FUNCTION_BLOCK basicEEEBruto (* Logica unica da elevatoria de esgoto bruto (3 bombas, 2 operando + 1 reserva) *)
  (* Standard: 61499-2 *)
  (* Version 1.6, 21/10/2026, Hidryco, Hidryco, 1.6: PID de nivel em Hz (minimo, maximo, preset e saida; 60 Hz = 100 %); STS_VELOCIDADE da IHM em Hz. 1.5: faixas da necessidade pela % da altura do poco (nivPct); stsNivel (IHM) continua em metros. 1.4: IHM: nivel, saida do PID, velocidade e tempo restante no maximo 1 vez por segundo (TICK). 1.3: pressao L/LL do PIT-01 inibida com as bombas paradas mesmo com cfgTempoPartidaPressao = 0. 1.2: emergencia do PCM NF. 1.1: emergencia do painel e falha de comunicacao dos ATV630. 1.0: faixas de nivel, revezamento por tempo, PID de velocidade, HH do Nereda, operacao pelas boias, falha de recalque *)
  PACKAGE Hidryco.HidrycoLib;
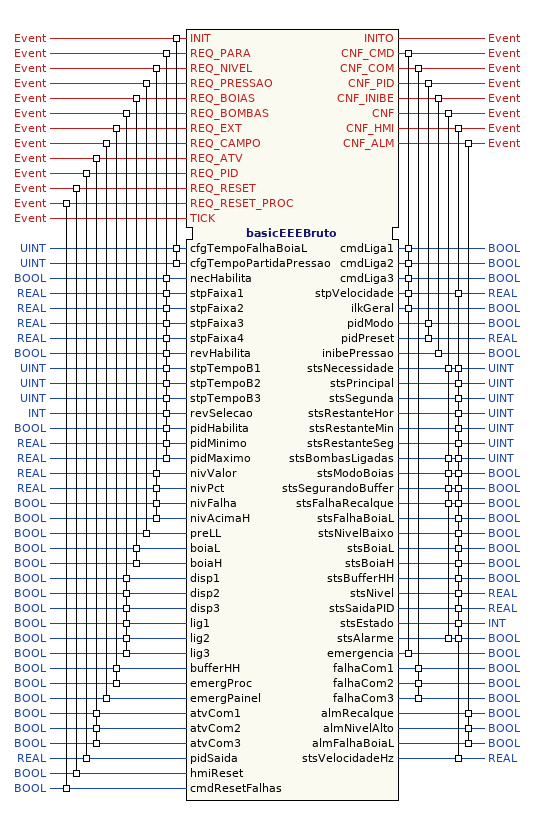
  EVENT_INPUT
    INIT WITH cfgTempoFalhaBoiaL, cfgTempoPartidaPressao; (* Inicializacao *)
    REQ_PARA WITH necHabilita, stpFaixa1, stpFaixa2, stpFaixa3, stpFaixa4, revHabilita, stpTempoB1, stpTempoB2, stpTempoB3, revSelecao, pidHabilita, pidMinimo, pidMaximo; (* Parametros da IHM (persistentes) *)
    REQ_NIVEL WITH nivValor, nivPct, nivFalha, nivAcimaH; (* LIT-03 *)
    REQ_PRESSAO WITH preLL; (* PIT-01 *)
    REQ_BOIAS WITH boiaL, boiaH; (* Boias *)
    REQ_BOMBAS WITH disp1, disp2, disp3, lig1, lig2, lig3; (* Estado das bombas *)
    REQ_EXT WITH bufferHH, emergProc; (* Processo *)
    REQ_CAMPO WITH emergPainel; (* Emergencia do painel *)
    REQ_ATV WITH atvCom1, atvCom2, atvCom3; (* Comunicacao dos ATV630 *)
    REQ_PID WITH pidSaida; (* Saida do PID *)
    REQ_RESET WITH hmiReset; (* Reset pela IHM *)
    REQ_RESET_PROC WITH cmdResetFalhas; (* Reset pelo processo *)
    TICK; (* Base de tempo de 1 s (E_CYCLE) *)
  END_EVENT
  EVENT_OUTPUT
    INITO; (* Inicializacao concluida *)
    CNF_CMD WITH cmdLiga1, cmdLiga2, cmdLiga3, stpVelocidade, ilkGeral, emergencia; (* Comandos para as bombas (na mudanca) *)
    CNF_COM WITH falhaCom1, falhaCom2, falhaCom3; (* Falha de comunicacao dos ATV630 para os motores (na mudanca e a cada leitura) *)
    CNF_PID WITH pidModo, pidPreset; (* Modo do pidCtl (na mudanca) *)
    CNF_INIBE WITH inibePressao; (* Inibicao dos alarmes baixos do PIT-01 (na mudanca) *)
    CNF WITH stsNecessidade, stsBombasLigadas, stsSegurandoBuffer, stsModoBoias, stsFalhaRecalque, stsAlarme; (* Status para o processo (na mudanca) *)
    CNF_HMI WITH stsNecessidade, stsPrincipal, stsSegunda, stsRestanteHor, stsRestanteMin, stsRestanteSeg, stsBombasLigadas, stsModoBoias, stsSegurandoBuffer, stsFalhaRecalque, stsFalhaBoiaL, stsNivelBaixo, stsBoiaL, stsBoiaH, stsBufferHH, stsNivel, stsSaidaPID, stpVelocidade, stsEstado, stsAlarme, stsVelocidadeHz; (* Status para a IHM (na mudanca) *)
    CNF_ALM WITH almRecalque, almNivelAlto, almFalhaBoiaL; (* Alarmes para os ALARM_BIT (na mudanca) *)
  END_EVENT
  VAR_INPUT
    cfgTempoFalhaBoiaL : UINT := 10; (* Operacao pelas boias com a boia LSL com defeito: bombas ficam ligadas este tempo (min) depois que a LSH desce *)
    cfgTempoPartidaPressao : UINT := 30; (* Alarmes L/LL do PIT-01 inibidos ate a bomba estar ligada ha este tempo (s); tambem inibidos com as bombas paradas *)
    necHabilita : BOOL; (* IHM: automatico da elevatoria habilitado (NEC_CMD_HABILITA) *)
    stpFaixa1 : REAL; (* IHM: com 1 bomba, desliga abaixo deste nivel (STP_LIMITE_FAIXA_1) *)
    stpFaixa2 : REAL; (* IHM: com 2 bombas, desliga a 2a abaixo deste nivel (STP_LIMITE_FAIXA_2) *)
    stpFaixa3 : REAL; (* IHM: parada, liga a 1a bomba neste nivel (STP_LIMITE_FAIXA_3) *)
    stpFaixa4 : REAL; (* IHM: com 1 bomba, liga a 2a neste nivel (STP_LIMITE_FAIXA_4) *)
    revHabilita : BOOL; (* IHM: revezamento por tempo habilitado (REV_CMD_HABILITA) *)
    stpTempoB1 : UINT; (* IHM: horas da bomba 1 como principal antes da troca; 0 = sem troca por tempo (STP_TEMPO_B1) *)
    stpTempoB2 : UINT; (* IHM: horas da bomba 2 como principal antes da troca; 0 = sem troca por tempo (STP_TEMPO_B2) *)
    stpTempoB3 : UINT; (* IHM: horas da bomba 3 como principal antes da troca; 0 = sem troca por tempo (STP_TEMPO_B3) *)
    revSelecao : INT; (* IHM: bomba principal 1, 2 ou 3 (CMD_SELECAO_BOMBA); comeca por ela ao escolher e a cada nova partida *)
    pidHabilita : BOOL; (* IHM: velocidade pelo PID de nivel (PID_CMD_HABILITA); FALSE = velocidade maxima *)
    pidMinimo : REAL; (* IHM: velocidade minima / saida minima do PID, % (STP_MINIMO) *)
    pidMaximo : REAL; (* IHM: velocidade maxima / saida maxima do PID, % (STP_MAXIMO) *)
    nivValor : REAL; (* LIT-03: nivel (unidade de engenharia) *)
    nivPct : REAL; (* LIT-03: nivel em % da altura do poco (faixas da necessidade) *)
    nivFalha : BOOL; (* LIT-03: sinal em falha agora *)
    nivAcimaH : BOOL; (* LIT-03: nivel acima do setpoint H agora (alarme H habilitado) *)
    preLL : BOOL; (* PIT-01: alarme LL de pressao (ja com o tempo do sensor) *)
    boiaL : BOOL; (* LSL-04: TRUE = boia levantada (nivel acima do baixo) *)
    boiaH : BOOL; (* LSH-05: TRUE = boia levantada (nivel alto) *)
    disp1 : BOOL; (* Bomba 1 disponivel para o automatico *)
    disp2 : BOOL; (* Bomba 2 disponivel para o automatico *)
    disp3 : BOOL; (* Bomba 3 disponivel para o automatico *)
    lig1 : BOOL; (* Bomba 1 ligada *)
    lig2 : BOOL; (* Bomba 2 ligada *)
    lig3 : BOOL; (* Bomba 3 ligada *)
    bufferHH : BOOL; (* Processo: nivel HH do tanque de equalizacao do Nereda (40-LT-0001) *)
    emergProc : BOOL; (* Processo: emergencia (entrada stsEmergencia do CAT) *)
    emergPainel : BOOL; (* Campo: emergencia do PCM EEE Bruto, NF (TRUE = normal; FALSE = em emergencia) *)
    atvCom1 : BOOL; (* ATV630 da bomba 1: comunicacao ativa (ComStatus do HW CAT) *)
    atvCom2 : BOOL; (* ATV630 da bomba 2: comunicacao ativa (ComStatus do HW CAT) *)
    atvCom3 : BOOL; (* ATV630 da bomba 3: comunicacao ativa (ComStatus do HW CAT) *)
    pidSaida : REAL; (* Saida do pidCtl (%) *)
    hmiReset : BOOL; (* IHM: reset *)
    cmdResetFalhas : BOOL; (* Processo: reset (com E_RESET_FALHAS) *)
  END_VAR
  VAR_OUTPUT
    cmdLiga1 : BOOL; (* Comando automatico da bomba 1 *)
    cmdLiga2 : BOOL; (* Comando automatico da bomba 2 *)
    cmdLiga3 : BOOL; (* Comando automatico da bomba 3 *)
    stpVelocidade : REAL; (* Velocidade das bombas ligadas (%) *)
    ilkGeral : BOOL; (* Intertravamento geral das bombas (LSL em nivel baixo ou falha de recalque); vale em qualquer modo *)
    pidModo : BOOL; (* pidCtl em automatico *)
    pidPreset : REAL; (* Valor do pidCtl em manual (%) *)
    inibePressao : BOOL; (* Inibe os alarmes L/LL do PIT-01 *)
    stsNecessidade : UINT; (* Numero de bombas pedidas (0, 1, 2) *)
    stsPrincipal : UINT; (* Bomba principal (1..3) *)
    stsSegunda : UINT; (* Bomba que entra como 2a (0 = nenhuma disponivel) *)
    stsRestanteHor : UINT; (* Tempo para a troca da principal (h) *)
    stsRestanteMin : UINT; (* Tempo para a troca da principal (min) *)
    stsRestanteSeg : UINT; (* Tempo para a troca da principal (s) *)
    stsBombasLigadas : UINT; (* Bombas ligadas *)
    stsModoBoias : BOOL; (* Operacao de emergencia pelas boias (LIT-03 em falha) *)
    stsSegurandoBuffer : BOOL; (* Elevatoria parada segurando o esgoto (HH do tanque do Nereda) *)
    stsFalhaRecalque : BOOL; (* Falha de recalque (pressao LL com bomba ligada) - memorizada ate o reset *)
    stsFalhaBoiaL : BOOL; (* Boia LSL com defeito (LSH levantada com a LSL abaixada) - memorizada ate o reset *)
    stsNivelBaixo : BOOL; (* LSL em nivel baixo: bombas intertravadas *)
    stsBoiaL : BOOL; (* LSL-04 *)
    stsBoiaH : BOOL; (* LSH-05 *)
    stsBufferHH : BOOL; (* HH do tanque do Nereda *)
    stsNivel : REAL; (* Nivel do poco *)
    stsSaidaPID : REAL; (* Saida do PID (%) *)
    stsEstado : INT; (* 0 parada, 1 bombeando, 2 segurando (HH Nereda), 3 pelas boias, 4 falha de recalque, 5 nivel baixo (LSL), 6 automatico desabilitado, 7 emergencia *)
    stsAlarme : BOOL; (* Algum alarme da elevatoria *)
    emergencia : BOOL; (* Emergencia para as bombas (painel OU processo) *)
    falhaCom1 : BOOL; (* Falha de comunicacao com o ATV630 da bomba 1 (publicada no stsFalhaComunicacao do motor) *)
    falhaCom2 : BOOL; (* Falha de comunicacao com o ATV630 da bomba 2 (publicada no stsFalhaComunicacao do motor) *)
    falhaCom3 : BOOL; (* Falha de comunicacao com o ATV630 da bomba 3 (publicada no stsFalhaComunicacao do motor) *)
    almRecalque : BOOL; (* ALARM_BIT falha de recalque *)
    almNivelAlto : BOOL; (* ALARM_BIT nivel alto (LSH) *)
    almFalhaBoiaL : BOOL; (* ALARM_BIT defeito da boia LSL *)
    stsVelocidadeHz : REAL; (* Velocidade enviada as bombas em Hz (IHM/SCADA) *)
  END_VAR
  VAR
    initDone : BOOL;
    initPass : BOOL;
    bReset : BOOL;
    bNivelRecebido : BOOL; (* Ja houve leitura do LIT-03 *)
    bBoiasRecebidas : BOOL; (* Ja houve leitura das boias *)
    bNivelOk : BOOL; (* LIT-03 valido *)
    bAlgumaLigada : BOOL;
    bLiberadoHH : BOOL; (* HH do Nereda: liberado pelo nivel H do poco *)
    iNec : UINT; (* Numero de bombas pedidas *)
    oldNec : UINT;
    bCampoRecebido : BOOL; (* Ja houve leitura da emergencia do painel *)
    iPrincipal : UINT := 1; (* Bomba principal (revezamento) *)
    iSel : INT; (* Selecao da principal valida (1..3) *)
    oldSel : INT; (* Ultima selecao aplicada *)
    iUso : UINT; (* Principal em uso (fixa indisponivel = proxima) *)
    iSeg : UINT; (* 2a bomba *)
    iProx : UINT;
    iCand : UINT;
    i : UINT;
    bDisp : BOOL;
    bDispP : BOOL;
    bLigP : BOOL;
    uSegPrincipal : UDINT; (* Segundos da principal ligada desde a ultima troca *)
    uLimite : UDINT;
    uResta : UDINT;
    uTempoBoia : UDINT; (* Contagem (s) da operacao pelas boias com a LSL com defeito *)
    uSegLigada : UDINT; (* Segundos com bomba ligada (inibicao do PIT-01) *)
    wCmd : WORD;
    oldCmd : WORD := 16#FFFF;
    oldVel : REAL := -1.0;
    oldPidModo : BOOL;
    oldPreset : REAL := -1.0;
    oldInibe : BOOL;
    wSts : WORD;
    oldSts : WORD := 16#FFFF;
    wHmi : WORD;
    oldHmi : WORD := 16#FFFF;
    oldNivel : REAL := -1.0;
    oldSaida : REAL := -1.0;
    oldResta : UDINT := 16#FFFFFFFF;
    hmiVel : REAL := -1.0;
    oldEstado : INT := -1;
    oldInfo : UINT := 16#FFFF;
    uInfo : UINT;
    wAlm : WORD;
    oldAlm : WORD := 16#FFFF;
    wCom : WORD;
    oldCom : WORD := 16#FFFF;
  END_VAR
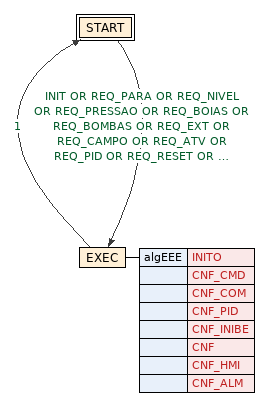
  EC_STATES
    START; (* Estado inicial *)
    EXEC : algEEE -> INITO, -> CNF_CMD, -> CNF_COM, -> CNF_PID, -> CNF_INIBE, -> CNF, -> CNF_HMI, -> CNF_ALM; (* Executa a logica; o algoritmo decide quais eventos saem *)
  END_STATES
  EC_TRANSITIONS
    START TO EXEC := INIT OR REQ_PARA OR REQ_NIVEL OR REQ_PRESSAO OR REQ_BOIAS OR REQ_BOMBAS OR REQ_EXT OR REQ_CAMPO OR REQ_ATV OR REQ_PID OR REQ_RESET OR REQ_RESET_PROC OR TICK;
    EXEC TO START := 1;
  END_TRANSITIONS
  ALGORITHM algEEE IN ST: (* Logica completa da elevatoria (um unico algoritmo) *)
(* =====================================================================
   basicEEEBruto v1.1 - Elevatoria de Esgoto Bruto (100-BS-01/02/03)
   Padrao das bibliotecas Schneider: eventos de saida desligados no inicio e
   ligados so na mudanca; tempos contados pelo TICK de 1 s (E_CYCLE do CAT).
   Regras (definidas pelo usuario, out/2026):
   - numero de bombas por faixas de nivel do LIT-03 (mesmas tags do CAT
     Necessidade_2_Equipamentos), no maximo 2; velocidade pelo PID de nivel;
   - revezamento: a principal selecionada (1, 2 ou 3) e a primeira a partir
     (ao escolher e sempre que as bombas partem de novo); com o revezamento
     habilitado troca apos STP_TEMPO_Bx horas ligada, na sequencia 1-2-3
     pulando a indisponivel; a 2a e a proxima da sequencia; principal
     indisponivel = troca na hora (tags do Revezamento_3_Motores);
   - HH do tanque do Nereda: a elevatoria para e segura o esgoto; volta a
     bombear quando o poco chega ao H dele (ou na LSH) - o tanque do Nereda
     tem extravasor; depois que esvazia ate a faixa 1, volta a segurar;
   - LIT-03 em falha: operacao pelas boias (LSH liga as 2 bombas na
     velocidade maxima; desligam quando a LSL abaixa; com a LSL com defeito,
     ficam cfgTempoFalhaBoiaL min depois que a LSH desce);
   - LSL abaixada desliga as bombas (ilkGeral) e elas voltam sozinhas;
   - PIT-01 em LL com bomba ligada = falha de recalque: para todas, alarma,
     memoriza ate o reset; L/LL do PIT-01 inibidos com as bombas paradas e
     nos primeiros cfgTempoPartidaPressao s depois da partida;
   - LSH so alarma (fora a operacao pelas boias e a liberacao do HH).
   v1.2: emergencia do PCM e NF (FALSE = em emergencia), so vale depois da
         1a leitura do campo.
   v1.1: emergencia do painel (campo) OU do processo vai para as bombas;
   falha de comunicacao de cada ATV630 = NOT ComStatus, publicada no
   stsFalhaComunicacao do motor (sem leitura = falha).
   ===================================================================== *)

(* ---- 0. Eventos de saida: so sai o que for ligado abaixo ---- *)
INITO     := FALSE;
CNF_CMD   := FALSE;
CNF_PID   := FALSE;
CNF_INIBE := FALSE;
CNF       := FALSE;
CNF_HMI   := FALSE;
CNF_ALM   := FALSE;
CNF_COM   := FALSE;

IF REQ_NIVEL THEN
    bNivelRecebido := TRUE;
END_IF;
IF REQ_BOIAS THEN
    bBoiasRecebidas := TRUE;
END_IF;
IF REQ_CAMPO THEN
    bCampoRecebido := TRUE;
END_IF;

(* ---- 1. Inicializacao ---- *)
IF INIT THEN
    initDone := TRUE;
    initPass := TRUE;
    INITO    := TRUE;
END_IF;
IF NOT initDone THEN
    RETURN;
END_IF;

bReset := (REQ_RESET AND hmiReset) OR (REQ_RESET_PROC AND cmdResetFalhas);
bAlgumaLigada := lig1 OR lig2 OR lig3;
stsBombasLigadas := 0;
IF lig1 THEN stsBombasLigadas := stsBombasLigadas + 1; END_IF;
IF lig2 THEN stsBombasLigadas := stsBombasLigadas + 1; END_IF;
IF lig3 THEN stsBombasLigadas := stsBombasLigadas + 1; END_IF;

(* ---- 2. Boias ---- *)
IF boiaH AND NOT boiaL THEN
    stsFalhaBoiaL := TRUE;                 (* LSH levantada com a LSL abaixada: LSL com defeito *)
END_IF;
IF bReset AND boiaL THEN
    stsFalhaBoiaL := FALSE;
END_IF;
(* nivel baixo: LSL abaixada (so se a LSL estiver confiavel); antes da 1a leitura, bloqueado *)
stsNivelBaixo := NOT bBoiasRecebidas OR (NOT boiaL AND NOT stsFalhaBoiaL);

(* ---- 3. Falha de recalque (PIT-01) ---- *)
IF bAlgumaLigada THEN
    IF TICK AND uSegLigada < UINT_TO_UDINT(cfgTempoPartidaPressao) THEN
        uSegLigada := uSegLigada + 1;
    END_IF;
ELSE
    uSegLigada := 0;
END_IF;
inibePressao := NOT bAlgumaLigada OR uSegLigada < UINT_TO_UDINT(cfgTempoPartidaPressao);   (* parada: inibido mesmo com o tempo = 0 *)
IF preLL AND NOT inibePressao THEN
    stsFalhaRecalque := TRUE;              (* pressao LL com bomba ligada: para todas *)
END_IF;
IF bReset AND NOT preLL THEN
    stsFalhaRecalque := FALSE;
END_IF;
ilkGeral := stsNivelBaixo OR stsFalhaRecalque;

(* ---- 3b. Emergencia e comunicacao dos ATV630 ---- *)
emergencia := emergProc OR (bCampoRecebido AND NOT emergPainel);   (* PCM: contato NF; sem leitura = sem emergencia *)
falhaCom1 := NOT atvCom1;
falhaCom2 := NOT atvCom2;
falhaCom3 := NOT atvCom3;

(* ---- 4. Origem do nivel ---- *)
bNivelOk := bNivelRecebido AND NOT nivFalha;
stsModoBoias := NOT bNivelOk;

(* ---- 5. HH do tanque do Nereda: segura enquanto o poco nao chega ao H ---- *)
IF NOT bufferHH THEN
    bLiberadoHH := FALSE;
ELSIF (bNivelOk AND nivAcimaH) OR boiaH THEN
    bLiberadoHH := TRUE;                   (* poco no H: volta a bombear (o Nereda tem extravasor) *)
END_IF;
stsSegurandoBuffer := necHabilita AND bufferHH AND NOT bLiberadoHH;

(* ---- 6. Numero de bombas ---- *)
IF NOT necHabilita OR stsSegurandoBuffer THEN
    iNec := 0;
    uTempoBoia := 0;
ELSIF NOT stsModoBoias THEN
    uTempoBoia := 0;
    IF iNec = 0 THEN
        IF nivPct >= stpFaixa3 THEN
            iNec := 1;
        END_IF;
    ELSIF iNec = 1 THEN
        IF nivPct >= stpFaixa4 THEN
            iNec := 2;
        ELSIF nivPct < stpFaixa1 THEN
            iNec := 0;
        END_IF;
    ELSE
        IF nivPct < stpFaixa2 THEN
            iNec := 1;
        END_IF;
    END_IF;
ELSE
    (* operacao de emergencia pelas boias *)
    IF boiaH THEN
        iNec := 2;
        uTempoBoia := UINT_TO_UDINT(cfgTempoFalhaBoiaL) * 60;
    ELSIF iNec > 0 THEN
        IF stsFalhaBoiaL THEN
            IF TICK AND uTempoBoia > 0 THEN
                uTempoBoia := uTempoBoia - 1;
            END_IF;
            IF uTempoBoia = 0 THEN
                iNec := 0;                 (* LSL com defeito: desliga pelo tempo *)
            END_IF;
        ELSIF NOT boiaL THEN
            iNec := 0;                     (* LSL abaixou *)
        END_IF;
    END_IF;
END_IF;
IF iNec = 0 AND oldNec > 0 THEN
    bLiberadoHH := FALSE;                  (* esvaziou: se o HH do Nereda continuar, volta a segurar *)
END_IF;
oldNec := iNec;
stsNecessidade := iNec;

(* ---- 7. Revezamento ---- *)
(* selecao da principal so 1, 2 ou 3 (0 gravado de antes vale 1); a selecionada vira a principal ao ser
   escolhida e sempre que as bombas partem de novo (todas paradas e sem necessidade); com o revezamento
   habilitado a troca por tempo segue a partir dela *)
iSel := revSelecao;
IF iSel < 1 OR iSel > 3 THEN
    iSel := 1;
END_IF;
IF iPrincipal < 1 OR iPrincipal > 3 THEN
    iPrincipal := INT_TO_UINT(iSel);
END_IF;
IF iSel <> oldSel THEN
    iPrincipal := INT_TO_UINT(iSel);
    uSegPrincipal := 0;
    oldSel := iSel;
END_IF;
IF iNec = 0 AND NOT lig1 AND NOT lig2 AND NOT lig3 THEN
    iPrincipal := INT_TO_UINT(iSel);       (* proxima partida comeca pela selecionada *)
    uSegPrincipal := 0;
END_IF;
(* proxima disponivel depois da principal, na sequencia 1-2-3 *)
iProx := 0;
iCand := iPrincipal;
FOR i := 1 TO 2 DO
    iCand := iCand + 1;
    IF iCand > 3 THEN
        iCand := 1;
    END_IF;
    IF iCand = 1 THEN
        bDisp := disp1;
    ELSIF iCand = 2 THEN
        bDisp := disp2;
    ELSE
        bDisp := disp3;
    END_IF;
    IF bDisp AND iProx = 0 THEN
        iProx := iCand;
    END_IF;
END_FOR;
IF iPrincipal = 1 THEN
    bDispP := disp1; bLigP := lig1;
ELSIF iPrincipal = 2 THEN
    bDispP := disp2; bLigP := lig2;
ELSE
    bDispP := disp3; bLigP := lig3;
END_IF;
IF revHabilita THEN
    IF NOT bDispP AND iProx <> 0 THEN
        iPrincipal := iProx;               (* principal indisponivel: troca na hora *)
        uSegPrincipal := 0;
    ELSE
        IF TICK AND bLigP AND uLimite > 0 THEN
            uSegPrincipal := uSegPrincipal + 1;
        END_IF;
        IF uLimite > 0 AND uSegPrincipal >= uLimite AND iProx <> 0 THEN
            iPrincipal := iProx;           (* venceu o tempo da principal *)
            uSegPrincipal := 0;
        END_IF;
    END_IF;
    iUso := iPrincipal;
ELSE
    (* sem revezamento: a selecionada e sempre a principal; indisponivel, a proxima assume so enquanto ela estiver fora *)
    IF NOT bDispP AND iProx <> 0 THEN
        iUso := iProx;
    ELSE
        iUso := iPrincipal;
    END_IF;
END_IF;
IF NOT revHabilita THEN
    uLimite := 0;
ELSIF iPrincipal = 1 THEN
    uLimite := UINT_TO_UDINT(stpTempoB1) * 3600;
ELSIF iPrincipal = 2 THEN
    uLimite := UINT_TO_UDINT(stpTempoB2) * 3600;
ELSE
    uLimite := UINT_TO_UDINT(stpTempoB3) * 3600;
END_IF;
(* 2a bomba: proxima disponivel depois da principal em uso *)
iSeg := 0;
iCand := iUso;
FOR i := 1 TO 2 DO
    iCand := iCand + 1;
    IF iCand > 3 THEN
        iCand := 1;
    END_IF;
    IF iCand = 1 THEN
        bDisp := disp1;
    ELSIF iCand = 2 THEN
        bDisp := disp2;
    ELSE
        bDisp := disp3;
    END_IF;
    IF bDisp AND iSeg = 0 THEN
        iSeg := iCand;
    END_IF;
END_FOR;
stsPrincipal := iUso;
stsSegunda := iSeg;
IF uLimite > uSegPrincipal THEN
    uResta := uLimite - uSegPrincipal;
ELSE
    uResta := 0;
END_IF;
stsRestanteHor := UDINT_TO_UINT(uResta / 3600);
stsRestanteMin := UDINT_TO_UINT((uResta MOD 3600) / 60);
stsRestanteSeg := UDINT_TO_UINT(uResta MOD 60);

(* ---- 8. Comandos ---- *)
cmdLiga1 := (iNec >= 1 AND iUso = 1) OR (iNec >= 2 AND iSeg = 1);
cmdLiga2 := (iNec >= 1 AND iUso = 2) OR (iNec >= 2 AND iSeg = 2);
cmdLiga3 := (iNec >= 1 AND iUso = 3) OR (iNec >= 2 AND iSeg = 3);

(* ---- 9. Velocidade ---- *)
pidModo := pidHabilita AND NOT stsModoBoias AND iNec > 0 AND bAlgumaLigada;
pidPreset := pidMinimo;
IF pidHabilita AND NOT stsModoBoias THEN
    IF pidModo THEN
        stpVelocidade := pidSaida / 0.6;   (* PID em Hz -> % das bombas *)
    ELSE
        stpVelocidade := pidMinimo / 0.6;        (* partida pela velocidade minima; o PID assume com a bomba ligada *)
    END_IF;
ELSE
    stpVelocidade := pidMaximo / 0.6;            (* PID desabilitado ou operacao pelas boias *)
END_IF;
stsSaidaPID := pidSaida;                   (* Hz *)
stsVelocidadeHz := stpVelocidade * 0.6;     (* IHM/SCADA em Hz *)

(* ---- 10. Status e alarmes ---- *)
stsBoiaL := boiaL;
stsBoiaH := boiaH;
stsBufferHH := bufferHH;
stsNivel := nivValor;
almRecalque := stsFalhaRecalque;
almNivelAlto := boiaH;
almFalhaBoiaL := stsFalhaBoiaL;
stsAlarme := almRecalque OR almNivelAlto OR almFalhaBoiaL;
IF emergencia THEN
    stsEstado := 7;
ELSIF stsFalhaRecalque THEN
    stsEstado := 4;
ELSIF stsNivelBaixo THEN
    stsEstado := 5;
ELSIF NOT necHabilita THEN
    stsEstado := 6;
ELSIF stsSegurandoBuffer THEN
    stsEstado := 2;
ELSIF stsModoBoias THEN
    stsEstado := 3;
ELSIF iNec > 0 THEN
    stsEstado := 1;
ELSE
    stsEstado := 0;
END_IF;

(* ---- 11. Eventos so na mudanca ---- *)
wCmd := 0;
IF cmdLiga1 THEN wCmd := wCmd OR 16#0001; END_IF;
IF cmdLiga2 THEN wCmd := wCmd OR 16#0002; END_IF;
IF cmdLiga3 THEN wCmd := wCmd OR 16#0004; END_IF;
IF ilkGeral THEN wCmd := wCmd OR 16#0008; END_IF;
IF emergencia THEN wCmd := wCmd OR 16#0010; END_IF;
CNF_CMD := initPass OR (wCmd <> oldCmd) OR (stpVelocidade <> oldVel);
CNF_PID := initPass OR (pidModo <> oldPidModo) OR (pidPreset <> oldPreset);
CNF_INIBE := initPass OR (inibePressao <> oldInibe);
wSts := 0;
IF stsSegurandoBuffer THEN wSts := wSts OR 16#0001; END_IF;
IF stsModoBoias       THEN wSts := wSts OR 16#0002; END_IF;
IF stsFalhaRecalque   THEN wSts := wSts OR 16#0004; END_IF;
IF stsAlarme          THEN wSts := wSts OR 16#0008; END_IF;
uInfo := iNec + stsBombasLigadas * 16 + iUso * 256 + iSeg * 4096;
CNF := initPass OR (wSts <> oldSts) OR (iNec <> (oldInfo MOD 16)) OR (stsBombasLigadas <> ((oldInfo / 16) MOD 16));
wHmi := wSts;
IF stsFalhaBoiaL  THEN wHmi := wHmi OR 16#0010; END_IF;
IF stsNivelBaixo  THEN wHmi := wHmi OR 16#0020; END_IF;
IF boiaL          THEN wHmi := wHmi OR 16#0040; END_IF;
IF boiaH          THEN wHmi := wHmi OR 16#0080; END_IF;
IF bufferHH       THEN wHmi := wHmi OR 16#0100; END_IF;
(* IHM: estado na hora; nivel, saida do PID, velocidade e tempo restante no maximo 1 vez por segundo (TICK) *)
CNF_HMI := initPass OR (wHmi <> oldHmi) OR (uInfo <> oldInfo) OR (stsEstado <> oldEstado)
           OR (TICK AND ((nivValor <> oldNivel) OR (pidSaida <> oldSaida) OR (stpVelocidade <> hmiVel) OR (uResta <> oldResta)));
wAlm := 0;
IF almRecalque   THEN wAlm := wAlm OR 16#0001; END_IF;
IF almNivelAlto  THEN wAlm := wAlm OR 16#0002; END_IF;
IF almFalhaBoiaL THEN wAlm := wAlm OR 16#0004; END_IF;
CNF_ALM := initPass OR (wAlm <> oldAlm);
wCom := 0;
IF falhaCom1 THEN wCom := wCom OR 16#0001; END_IF;
IF falhaCom2 THEN wCom := wCom OR 16#0002; END_IF;
IF falhaCom3 THEN wCom := wCom OR 16#0004; END_IF;
CNF_COM := initPass OR REQ_ATV OR (wCom <> oldCom);   (* a cada leitura: tambem republica depois do INIT do publicador *)
oldCmd := wCmd;
oldVel := stpVelocidade;
oldPidModo := pidModo;
oldPreset := pidPreset;
oldInibe := inibePressao;
oldSts := wSts;
oldHmi := wHmi;
oldInfo := uInfo;
oldEstado := stsEstado;
IF CNF_HMI THEN
    oldNivel := nivValor; oldSaida := pidSaida; oldResta := uResta; hmiVel := stpVelocidade;
END_IF;
oldAlm := wAlm;
oldCom := wCom;

initPass := FALSE;
  END_ALGORITHM
END_FUNCTION_BLOCK
